(* Logix 5000 project; controller SmartManufacturingCell Emulate 5570 rev 33.11; software revision 33.03; part 3 of 5 *)
(* tags used below, declared in another part *)
   ClearCell_CommandsReleased : BOOL;
   ClearCell_EquipmentReady : BOOL;
   ClearCellRequestONS : BOOL;
   Exit_ReadyForIndex : BOOL;
   Filling_ReadyForIndex : BOOL;
   Index_CommandsReleased : BOOL;
   Index_EquipmentReady : BOOL;
   IndexConfirmTimeout : TIMER;   // Non-retentive timer; preset in milliseconds.
   IndexTimeout : TIMER;   // Non-retentive timer; preset in milliseconds.
   Inspection_ReadyForIndex : BOOL;
   Production_CycleHealthy : BOOL;
   Production_ResetAllowed : BOOL;
   Production_ResetCommandsReleased : BOOL;
   Production_SensorsClear : BOOL;
   Production_TrackingEmpty : BOOL;
   ProductionResetONS : BOOL;
   TrackingMismatchDelay : TIMER;   // Non-retentive timer; preset in milliseconds.
   Conveyor_Flt_FailToStart : BOOL;   // Conveyor commanded but running feedback missing for 2 s Latched; clear cell, remove cause, then fresh Reset.
   Exit_Flt_DischargeTimeout : BOOL;   // Good or reject bottle departure not confirmed within 3 s Latched; clear cell, remove cause, then fresh Reset.
   Exit_Sts_State : DINT;   // 0 Empty; 10 Waiting; 20 Good discharge; 30 Extending; 40 Reject discharge; 50 Retracting; 60 Complete; 90 Faulted
   Filling_Flt_FillTimeout : BOOL;   // Fill completion not received within 4 s Latched; clear cell, remove cause, then fresh Reset.
   Filling_Flt_ValveFailToClose : BOOL;   // Fill valve did not close within 2 s Latched; clear cell, remove cause, then fresh Reset.
   Filling_Sts_State : DINT;   // 0 Empty; 10 Waiting; 20 Filling; 30 Closing; 40 Complete; 90 Faulted
   HMI_Cmd_ClearCell : BOOL;   // Request removal of simulated bottles during fault recovery
   HMI_Cmd_ConveyorJog : BOOL;   // Request conveyor movement while held
   HMI_Cmd_FillValveOpen : BOOL;
   HMI_Cmd_LoadBottle : BOOL;   // Request one simulated bottle at the available entry position
   HMI_Cmd_RejectExtend : BOOL;
   HMI_Cmd_Reset : BOOL;   // Request fault reset after recovery conditions are satisfied
   HMI_Cmd_Start : BOOL;   // Request automatic production start
   HMI_Cmd_Stop : BOOL;   // Request controlled production stop
   Inspection_Flt_Timeout : BOOL;   // Inspection did not finish within 3 s Latched; clear cell, remove cause, then fresh Reset.
   Inspection_Sts_State : DINT;   // 0 Empty; 10 Waiting; 20 Inspecting; 40 Complete; 90 Faulted
   Production_Bottles : UDT_Bottle[4];
   Production_Flt_IndexConfirmTimeout : BOOL;   // Post-index positions not confirmed within 1 s Latched; clear cell, remove cause, then fresh Reset.
   Production_Flt_IndexInterlock : BOOL;   // Movement interlock lost during indexing Latched; clear cell, remove cause, then fresh Reset.
   Production_Flt_IndexTimeout : BOOL;   // Index completion not received within 3 s Latched; clear cell, remove cause, then fresh Reset.
   Production_Flt_InvalidConfiguration : BOOL;   // Fill or inspection time outside permitted limits Latched; clear cell, remove cause, then fresh Reset.
   Production_Flt_InvalidState : BOOL;   // Machine, sequence, station state, or mode combination invalid Latched; clear cell, remove cause, then fresh Reset.
   Production_Flt_StartupRecoveryRequired : BOOL;   // Restart found bottles or interrupted activity Latched; clear cell, remove cause, then fresh Reset.
   Production_Flt_TrackingMismatch : BOOL;   // Stationary bottle tracking and sensors disagree or processing history invalid Latched; clear cell, remove cause, then fr
   Production_Stats_RecoveryLossCount : DINT;   // Retained RecoveryLossCount; count only confirmed departures (recovery losses separate).
   Production_Sts_ClearCellAccepted : BOOL;
   Production_Sts_ClearCellAllowed : BOOL;
   Production_Sts_IndexAllowed : BOOL;
   Production_Sts_IndexCommitted : BOOL;   // Bottle records transferred for the current confirmed index; cleared outside ConfirmPositions.
   Production_Sts_IndexDemand : BOOL;
   Production_Sts_IndexPositionsMatch : BOOL;   // Post-index positions verified in ConfirmPositions with conveyor stopped.
   Production_Sts_LoadAccepted : BOOL;
   Production_Sts_ResetAccepted : BOOL;
   Production_Sts_SequenceState : DINT;   // 0 = Idle 10 = ProcessStations 20 = Indexing 30 = ConfirmPositions
   Production_Sts_StationsReady : BOOL;
   Reject_Flt_FailToExtend : BOOL;   // Reject actuator did not extend within 2 s Latched; clear cell, remove cause, then fresh Reset.
   Reject_Flt_FailToRetract : BOOL;   // Reject actuator did not retract within 2 s Latched; clear cell, remove cause, then fresh Reset.
   Sim_In_ConveyorRunning : BOOL;   // Simulated conveyor movement feedback
   Sim_In_EntryPE : BOOL;   // Simulated bottle detected at entry
   Sim_In_ExitPE : BOOL;   // Simulated bottle detected at Reject/Exit position
   Sim_In_FillPE : BOOL;   // Simulated bottle detected at filling position
   Sim_In_FillValveClosed : BOOL;   // Simulated fill valve confirmed closed
   Sim_In_GoodExitPE : BOOL;   // Bottle detected passing through good discharge path
   Sim_In_IndexComplete : BOOL;   // Simulated conveyor completed one station-spacing movement
   Sim_In_InspectionPE : BOOL;   // Simulated bottle detected at inspection position
   Sim_In_RejectExitPE : BOOL;   // Bottle detected passing through reject discharge path
   Sim_In_RejectExtended : BOOL;   // Simulated reject actuator confirmed extended
   Sim_In_RejectRetracted : BOOL;   // Simulated reject actuator confirmed retracted
   Sim_Out_ConveyorRun : BOOL;   // Command simulated conveyor to run
   Sim_Out_FillValveOpen : BOOL;   // Command simulated fill valve to open
   Sim_Out_GoodDischargeRun : BOOL;   // Command simulated good-bottle discharge mechanism to run
   Sim_Out_RejectExtend : BOOL;   // Command simulated reject actuator to extend
   Sys_Sts_AutoMode : BOOL;   // Auto mode accepted and active
   Sys_Sts_BlockingFault : BOOL;   // Active blocking fault prevents production and manual equipment operation.
   Sys_Sts_MachineState : DINT;   // 0 = Stopped 10 = Running 20 = Stopping 30 = Faulted
   Sys_Sts_ManualMode : BOOL;   // Manual mode accepted and active
   Sys_Sts_ResetAllowed : BOOL;   // Sys Sts ResetAllowed
   Sys_Sts_StartupReady : BOOL;   // Sys Sts StartupReady
(* Program_Production, continued *)

ROUTINE Bottle_Tracking   (* structured text *)
   if Production_Sts_SequenceState <> 30 then
   	Production_Sts_IndexCommitted := 0;
   elsif Production_Sts_IndexPositionsMatch AND NOT Production_Sts_IndexCommitted then
   
   	// Copy downstream first to preserve seach source record.
   	COP(Production_Bottles[2], Production_Bottles[3], 1);
   	COP(Production_Bottles[1], Production_Bottles[2], 1);
   	COP(Production_Bottles[0], Production_Bottles[1], 1);
   
    	// Entry is empty after the confirmed movement.
       Production_Bottles[0].Occupied := 0;
       Production_Bottles[0].FillComplete := 0;
       Production_Bottles[0].InspectionComplete := 0;
       Production_Bottles[0].RejectRequired := 0;
   
       Production_Sts_IndexCommitted := 1;
   end_if;
END_ROUTINE

ROUTINE Clear_Cell   (* ladder *)
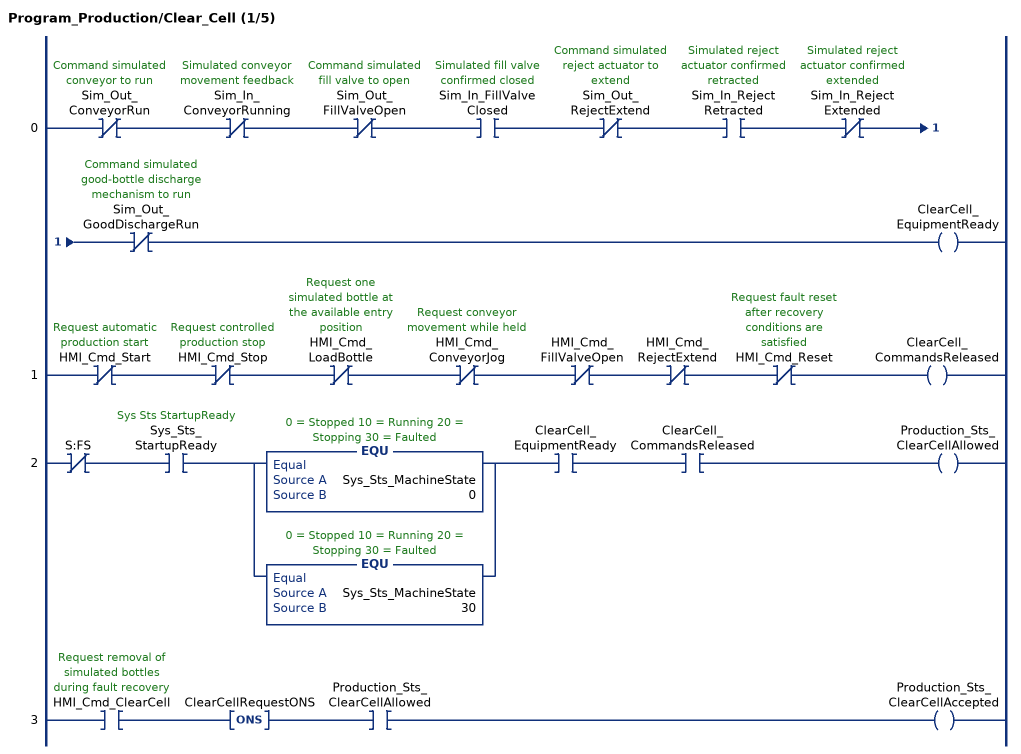
   0: XIO(Sim_Out_ConveyorRun)XIO(Sim_In_ConveyorRunning)XIO(Sim_Out_FillValveOpen)XIC(Sim_In_FillValveClosed)XIO(Sim_Out_RejectExtend)XIC(Sim_In_RejectRetracted)XIO(Sim_In_RejectExtended)XIO(Sim_Out_GoodDischargeRun)OTE(ClearCell_EquipmentReady);
   1: XIO(HMI_Cmd_Start)XIO(HMI_Cmd_Stop)XIO(HMI_Cmd_LoadBottle)XIO(HMI_Cmd_ConveyorJog)XIO(HMI_Cmd_FillValveOpen)XIO(HMI_Cmd_RejectExtend)XIO(HMI_Cmd_Reset)OTE(ClearCell_CommandsReleased);
   2: XIO(S:FS)XIC(Sys_Sts_StartupReady)[EQU(Sys_Sts_MachineState,0) ,EQU(Sys_Sts_MachineState,30) ]XIC(ClearCell_EquipmentReady)XIC(ClearCell_CommandsReleased)OTE(Production_Sts_ClearCellAllowed);
   3: XIC(HMI_Cmd_ClearCell)ONS(ClearCellRequestONS)XIC(Production_Sts_ClearCellAllowed)OTE(Production_Sts_ClearCellAccepted);
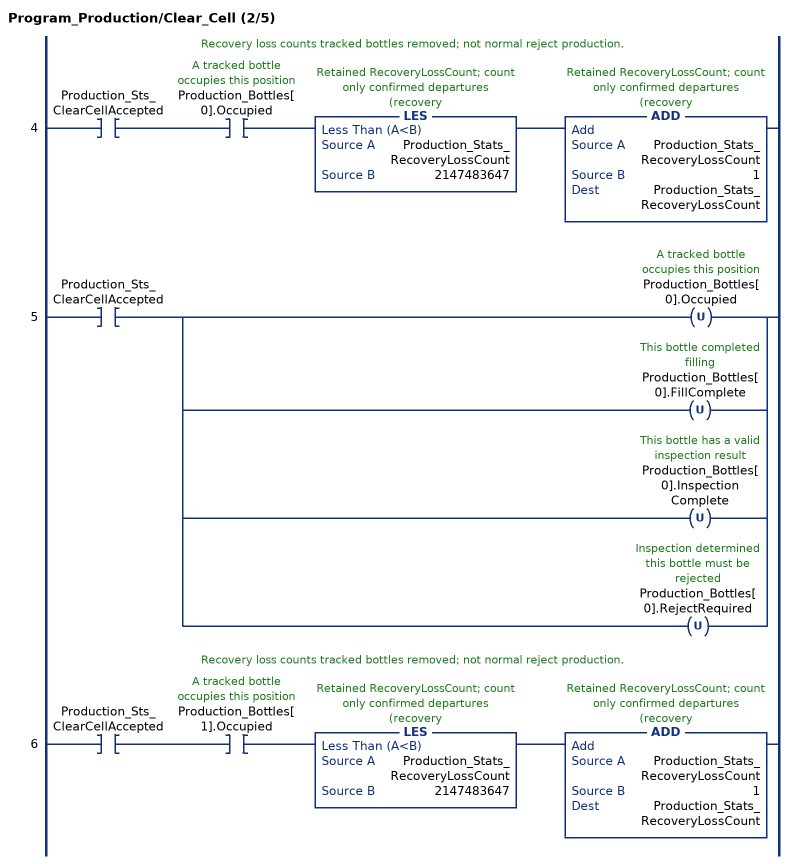
   // Recovery loss counts tracked bottles removed; not normal reject production.
   4: XIC(Production_Sts_ClearCellAccepted)XIC(Production_Bottles[0].Occupied)LES(Production_Stats_RecoveryLossCount,2147483647)ADD(Production_Stats_RecoveryLossCount,1,Production_Stats_RecoveryLossCount);
   5: XIC(Production_Sts_ClearCellAccepted)[OTU(Production_Bottles[0].Occupied) ,OTU(Production_Bottles[0].FillComplete) ,OTU(Production_Bottles[0].InspectionComplete) ,OTU(Production_Bottles[0].RejectRequired) ];
   // Recovery loss counts tracked bottles removed; not normal reject production.
   6: XIC(Production_Sts_ClearCellAccepted)XIC(Production_Bottles[1].Occupied)LES(Production_Stats_RecoveryLossCount,2147483647)ADD(Production_Stats_RecoveryLossCount,1,Production_Stats_RecoveryLossCount);
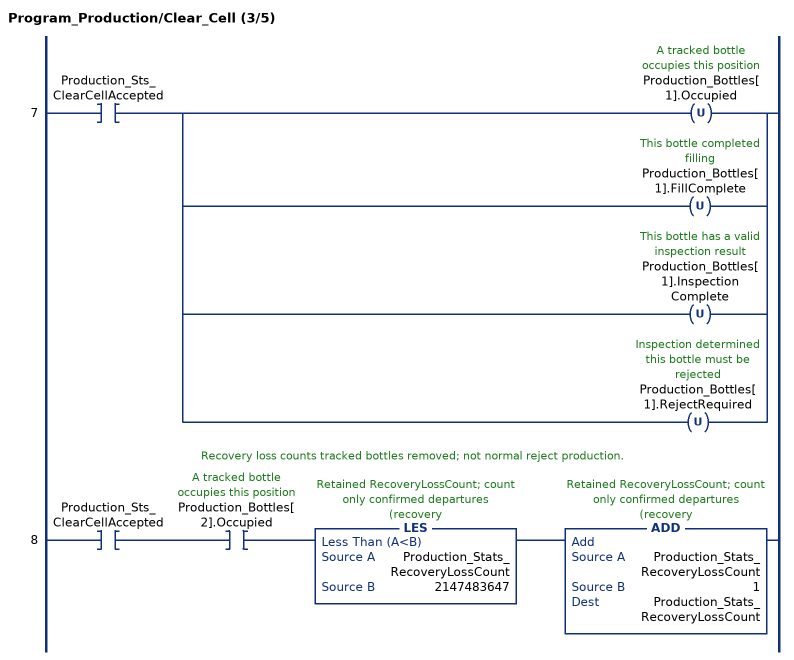
   7: XIC(Production_Sts_ClearCellAccepted)[OTU(Production_Bottles[1].Occupied) ,OTU(Production_Bottles[1].FillComplete) ,OTU(Production_Bottles[1].InspectionComplete) ,OTU(Production_Bottles[1].RejectRequired) ];
   // Recovery loss counts tracked bottles removed; not normal reject production.
   8: XIC(Production_Sts_ClearCellAccepted)XIC(Production_Bottles[2].Occupied)LES(Production_Stats_RecoveryLossCount,2147483647)ADD(Production_Stats_RecoveryLossCount,1,Production_Stats_RecoveryLossCount);
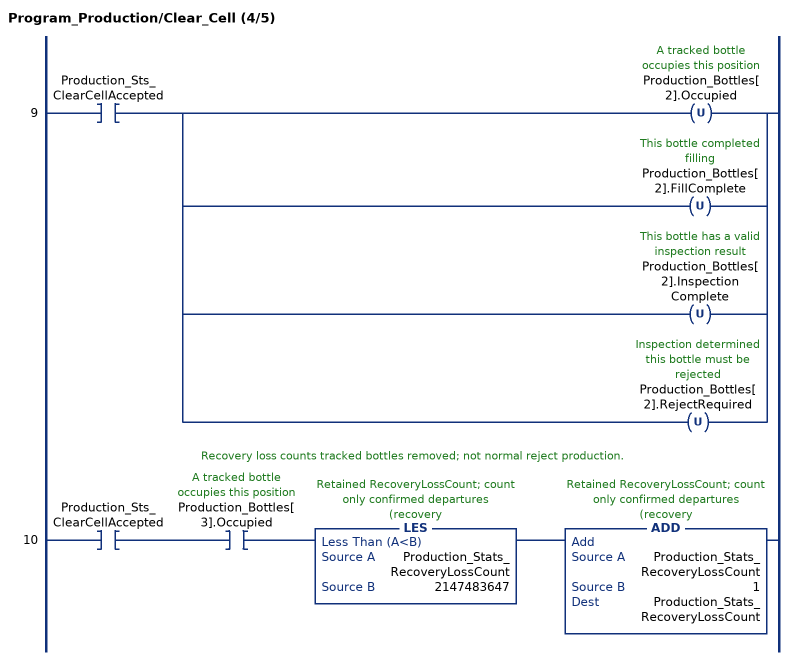
   9: XIC(Production_Sts_ClearCellAccepted)[OTU(Production_Bottles[2].Occupied) ,OTU(Production_Bottles[2].FillComplete) ,OTU(Production_Bottles[2].InspectionComplete) ,OTU(Production_Bottles[2].RejectRequired) ];
   // Recovery loss counts tracked bottles removed; not normal reject production.
   10: XIC(Production_Sts_ClearCellAccepted)XIC(Production_Bottles[3].Occupied)LES(Production_Stats_RecoveryLossCount,2147483647)ADD(Production_Stats_RecoveryLossCount,1,Production_Stats_RecoveryLossCount);
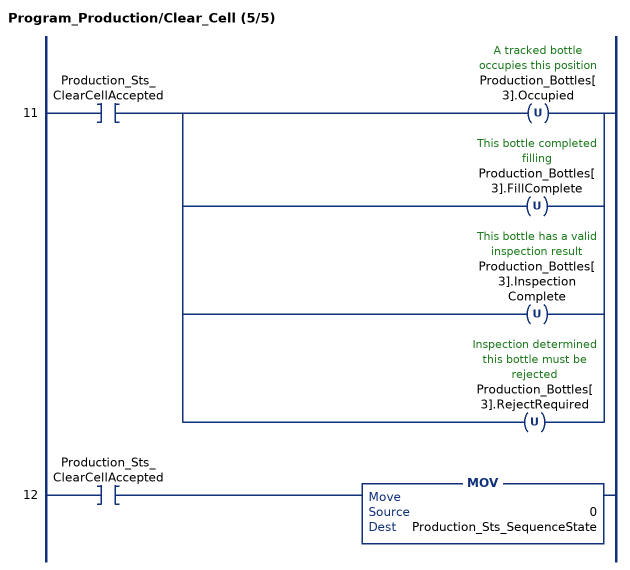
   11: XIC(Production_Sts_ClearCellAccepted)[OTU(Production_Bottles[3].Occupied) ,OTU(Production_Bottles[3].FillComplete) ,OTU(Production_Bottles[3].InspectionComplete) ,OTU(Production_Bottles[3].RejectRequired) ];
   12: XIC(Production_Sts_ClearCellAccepted)MOV(0,Production_Sts_SequenceState);
END_ROUTINE

ROUTINE Index_Confirmation   (* structured text *)
   Production_Sts_IndexPositionsMatch :=
       (Production_Sts_SequenceState = 30)
       AND (
           (Sys_Sts_MachineState = 10)
           OR (Sys_Sts_MachineState = 20)
       )
       AND Sys_Sts_AutoMode
       AND NOT Sys_Sts_ManualMode
       AND NOT Sys_Sts_BlockingFault
       AND NOT Sim_Out_ConveyorRun
       AND NOT Sim_In_ConveyorRunning
       AND NOT Production_Bottles[3].Occupied
       AND NOT Sim_In_EntryPE
       AND NOT (Sim_In_FillPE XOR Production_Bottles[0].Occupied)
       AND NOT (Sim_In_InspectionPE XOR Production_Bottles[1].Occupied)
       AND NOT (Sim_In_ExitPE XOR Production_Bottles[2].Occupied);
END_ROUTINE

ROUTINE Index_Permissives   (* ladder *)
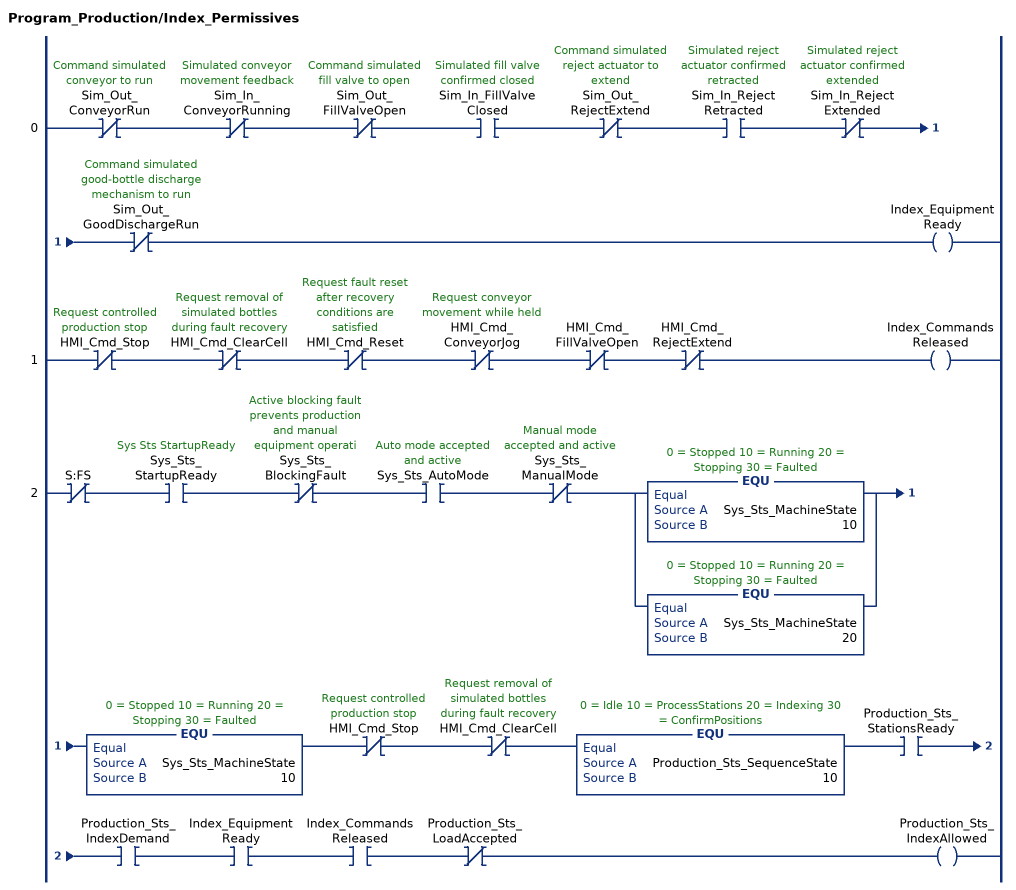
   0: XIO(Sim_Out_ConveyorRun)XIO(Sim_In_ConveyorRunning)XIO(Sim_Out_FillValveOpen)XIC(Sim_In_FillValveClosed)XIO(Sim_Out_RejectExtend)XIC(Sim_In_RejectRetracted)XIO(Sim_In_RejectExtended)XIO(Sim_Out_GoodDischargeRun)OTE(Index_EquipmentReady);
   1: XIO(HMI_Cmd_Stop)XIO(HMI_Cmd_ClearCell)XIO(HMI_Cmd_Reset)XIO(HMI_Cmd_ConveyorJog)XIO(HMI_Cmd_FillValveOpen)XIO(HMI_Cmd_RejectExtend)OTE(Index_CommandsReleased);
   2: XIO(S:FS)XIC(Sys_Sts_StartupReady)XIO(Sys_Sts_BlockingFault)XIC(Sys_Sts_AutoMode)XIO(Sys_Sts_ManualMode)[EQU(Sys_Sts_MachineState,10) ,EQU(Sys_Sts_MachineState,20) ]EQU(Sys_Sts_MachineState,10)XIO(HMI_Cmd_Stop)XIO(HMI_Cmd_ClearCell)EQU(Production_Sts_SequenceState,10)XIC(Production_Sts_StationsReady)XIC(Production_Sts_IndexDemand)XIC(Index_EquipmentReady)XIC(Index_CommandsReleased)XIO(Production_Sts_LoadAccepted)OTE(Production_Sts_IndexAllowed);
END_ROUTINE

ROUTINE Index_Readiness   (* ladder *)
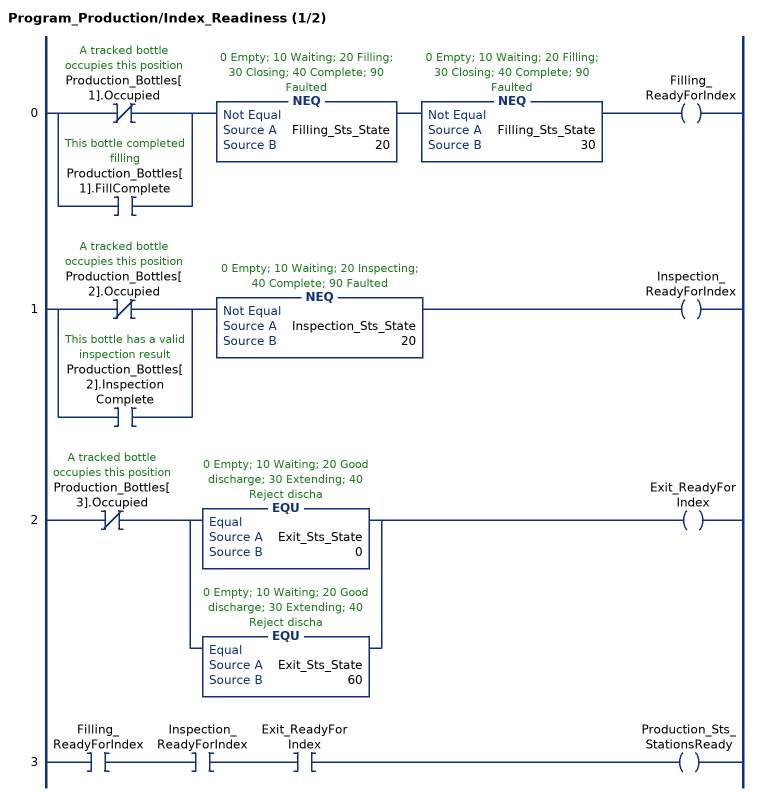
   0: [XIO(Production_Bottles[1].Occupied) ,XIC(Production_Bottles[1].FillComplete) ]NEQ(Filling_Sts_State,20)NEQ(Filling_Sts_State,30)OTE(Filling_ReadyForIndex);
   1: [XIO(Production_Bottles[2].Occupied) ,XIC(Production_Bottles[2].InspectionComplete) ]NEQ(Inspection_Sts_State,20)OTE(Inspection_ReadyForIndex);
   2: XIO(Production_Bottles[3].Occupied)[EQU(Exit_Sts_State,0) ,EQU(Exit_Sts_State,60) ]OTE(Exit_ReadyForIndex);
   3: XIC(Filling_ReadyForIndex)XIC(Inspection_ReadyForIndex)XIC(Exit_ReadyForIndex)OTE(Production_Sts_StationsReady);
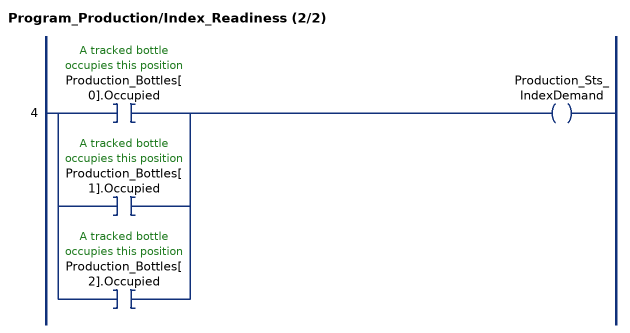
   4: [XIC(Production_Bottles[0].Occupied) ,XIC(Production_Bottles[1].Occupied) ,XIC(Production_Bottles[2].Occupied) ]OTE(Production_Sts_IndexDemand);
END_ROUTINE

ROUTINE MainRoutine   (* ladder *)
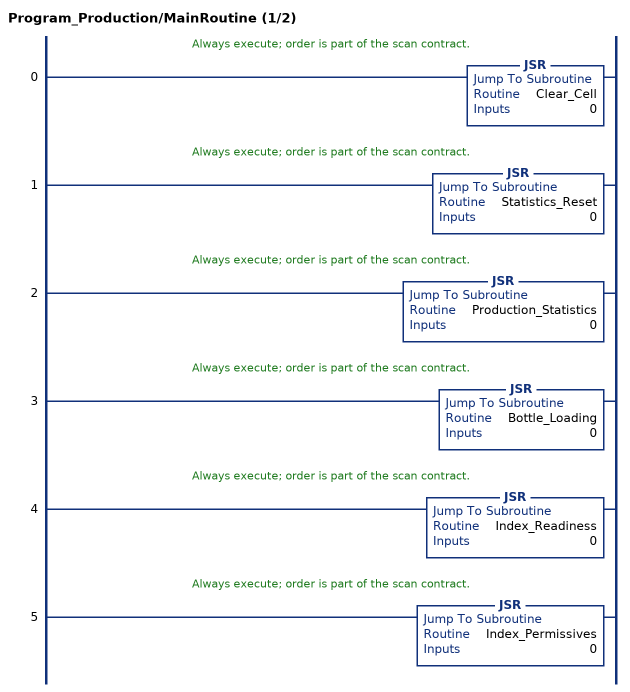
   // Always execute; order is part of the scan contract.
   0: JSR(Clear_Cell,0);
   // Always execute; order is part of the scan contract.
   1: JSR(Statistics_Reset,0);
   // Always execute; order is part of the scan contract.
   2: JSR(Production_Statistics,0);
   // Always execute; order is part of the scan contract.
   3: JSR(Bottle_Loading,0);
   // Always execute; order is part of the scan contract.
   4: JSR(Index_Readiness,0);
   // Always execute; order is part of the scan contract.
   5: JSR(Index_Permissives,0);
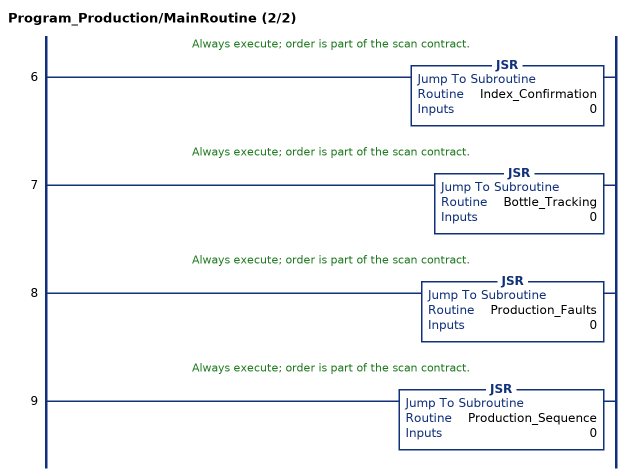
   // Always execute; order is part of the scan contract.
   6: JSR(Index_Confirmation,0);
   // Always execute; order is part of the scan contract.
   7: JSR(Bottle_Tracking,0);
   // Always execute; order is part of the scan contract.
   8: JSR(Production_Faults,0);
   // Always execute; order is part of the scan contract.
   9: JSR(Production_Sequence,0);
END_ROUTINE

ROUTINE Production_Faults   (* ladder *)
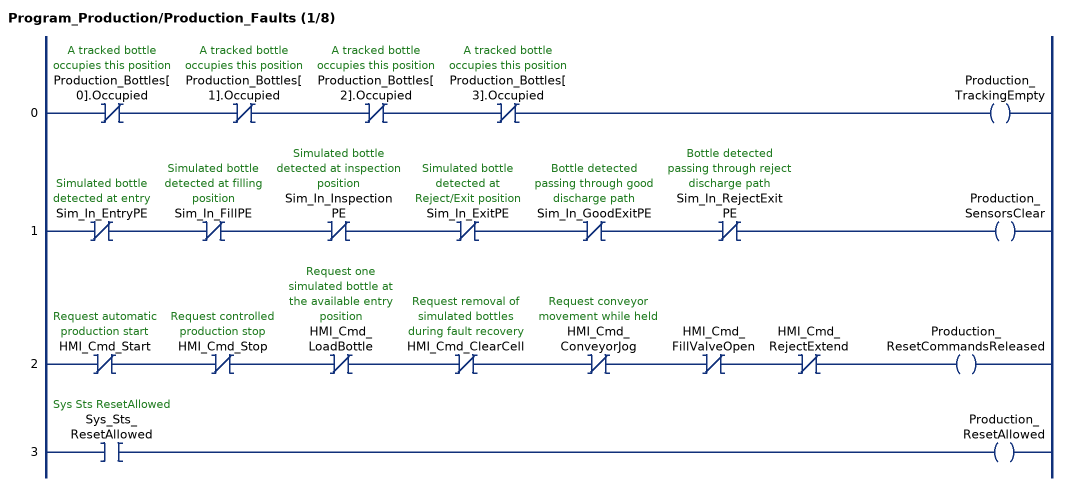
   0: XIO(Production_Bottles[0].Occupied)XIO(Production_Bottles[1].Occupied)XIO(Production_Bottles[2].Occupied)XIO(Production_Bottles[3].Occupied)OTE(Production_TrackingEmpty);
   1: XIO(Sim_In_EntryPE)XIO(Sim_In_FillPE)XIO(Sim_In_InspectionPE)XIO(Sim_In_ExitPE)XIO(Sim_In_GoodExitPE)XIO(Sim_In_RejectExitPE)OTE(Production_SensorsClear);
   2: XIO(HMI_Cmd_Start)XIO(HMI_Cmd_Stop)XIO(HMI_Cmd_LoadBottle)XIO(HMI_Cmd_ClearCell)XIO(HMI_Cmd_ConveyorJog)XIO(HMI_Cmd_FillValveOpen)XIO(HMI_Cmd_RejectExtend)OTE(Production_ResetCommandsReleased);
   3: XIC(Sys_Sts_ResetAllowed)OTE(Production_ResetAllowed);
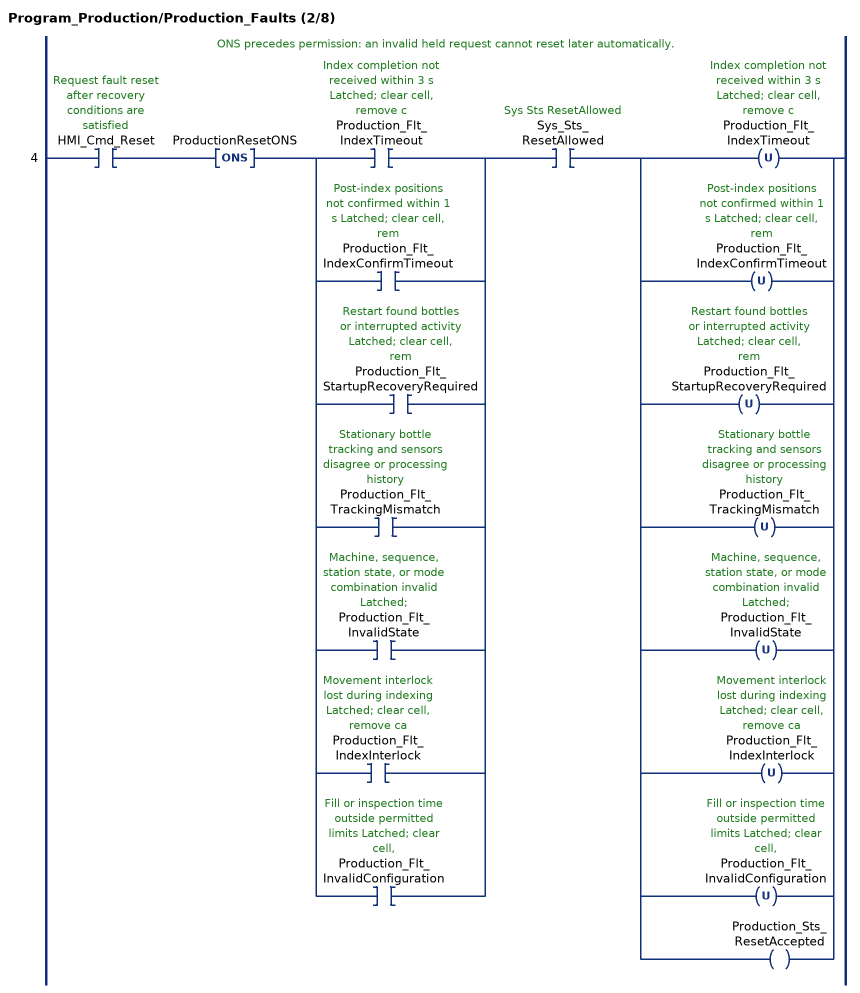
   // ONS precedes permission: an invalid held request cannot reset later automatically.
   4: XIC(HMI_Cmd_Reset)ONS(ProductionResetONS)[XIC(Production_Flt_IndexTimeout) ,XIC(Production_Flt_IndexConfirmTimeout) ,XIC(Production_Flt_StartupRecoveryRequired) ,XIC(Production_Flt_TrackingMismatch) ,XIC(Production_Flt_InvalidState) ,XIC(Production_Flt_IndexInterlock) ,XIC(Production_Flt_InvalidConfiguration) ]XIC(Sys_Sts_ResetAllowed)[OTU(Production_Flt_IndexTimeout) ,OTU(Production_Flt_IndexConfirmTimeout) ,OTU(Production_Flt_StartupRecoveryRequired) ,OTU(Production_Flt_TrackingMismatch) ,OTU(Production_Flt_InvalidState) ,OTU(Production_Flt_IndexInterlock) ,OTU(Production_Flt_InvalidConfiguration) ,OTE(Production_Sts_ResetAccepted) ];
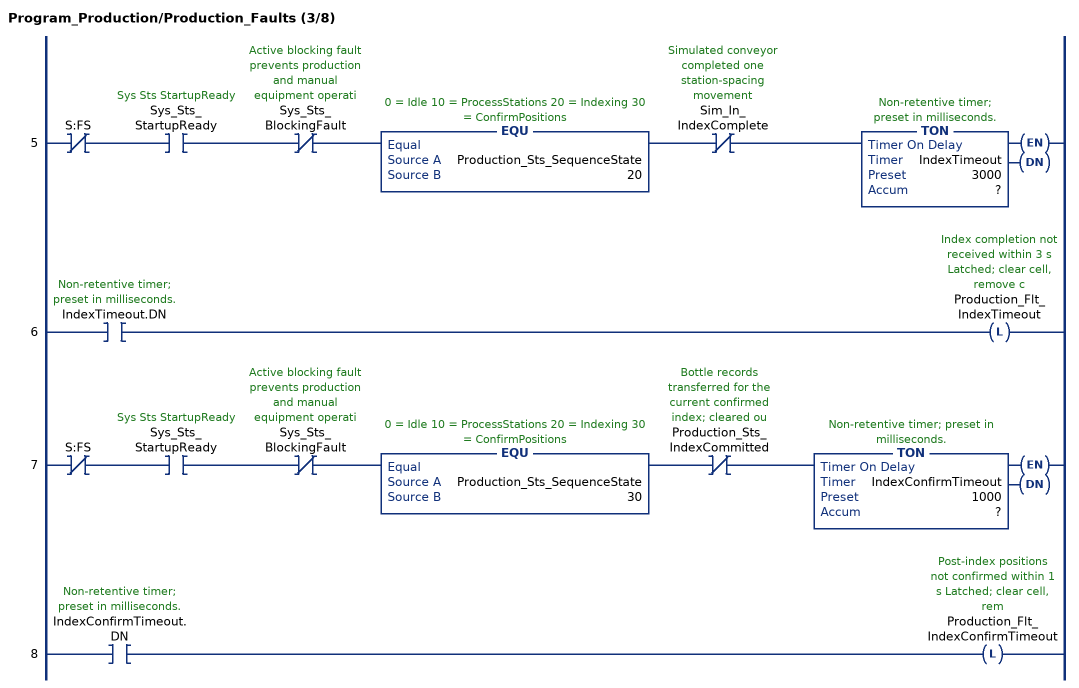
   5: XIO(S:FS)XIC(Sys_Sts_StartupReady)XIO(Sys_Sts_BlockingFault)EQU(Production_Sts_SequenceState,20)XIO(Sim_In_IndexComplete)TON(IndexTimeout,?,?);
   6: XIC(IndexTimeout.DN)OTL(Production_Flt_IndexTimeout);
   7: XIO(S:FS)XIC(Sys_Sts_StartupReady)XIO(Sys_Sts_BlockingFault)EQU(Production_Sts_SequenceState,30)XIO(Production_Sts_IndexCommitted)TON(IndexConfirmTimeout,?,?);
   8: XIC(IndexConfirmTimeout.DN)OTL(Production_Flt_IndexConfirmTimeout);
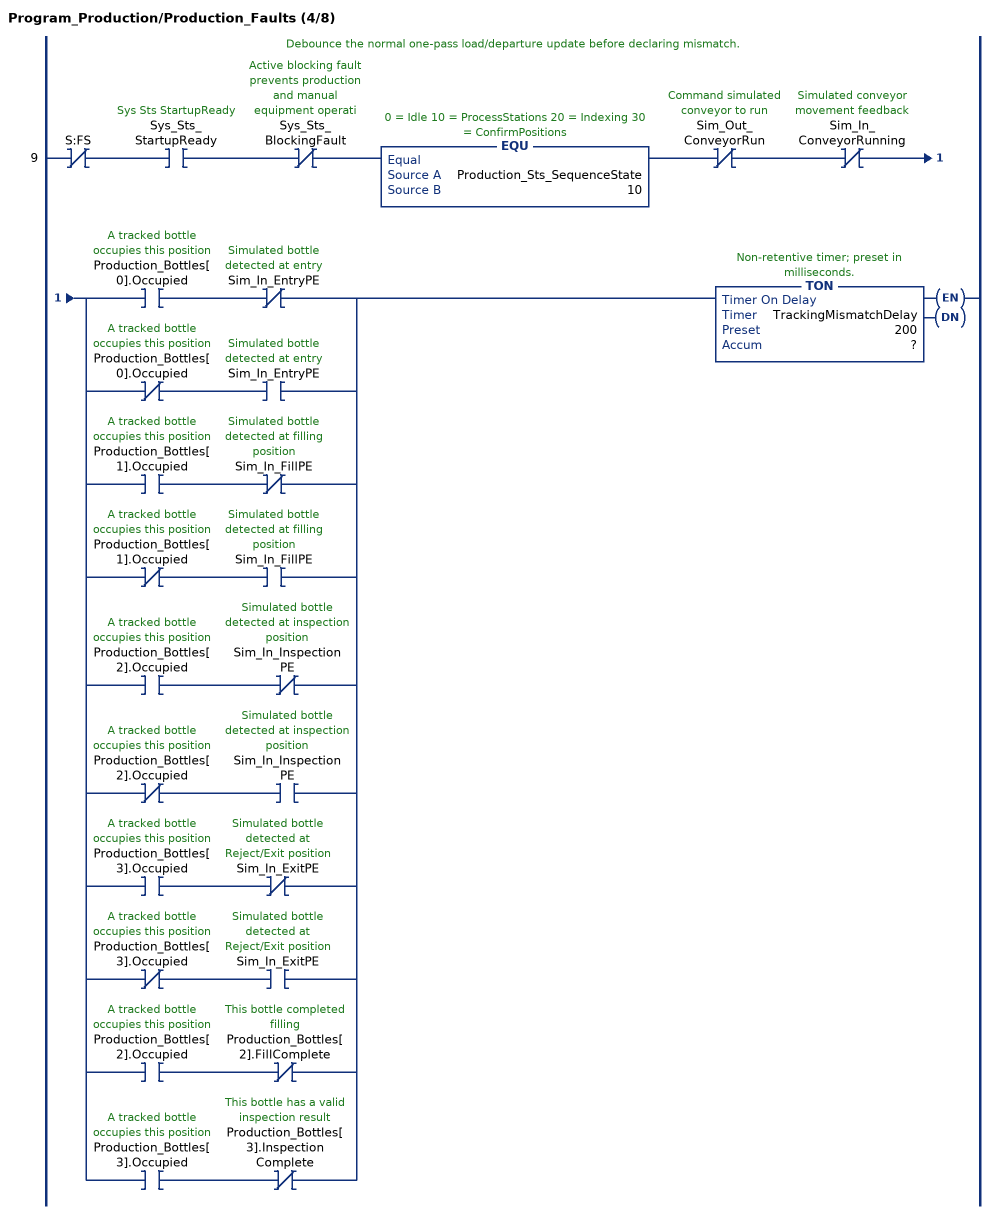
   // Debounce the normal one-pass load/departure update before declaring mismatch.
   9: XIO(S:FS)XIC(Sys_Sts_StartupReady)XIO(Sys_Sts_BlockingFault)EQU(Production_Sts_SequenceState,10)XIO(Sim_Out_ConveyorRun)XIO(Sim_In_ConveyorRunning)[[XIC(Production_Bottles[0].Occupied) XIO(Sim_In_EntryPE) ,XIO(Production_Bottles[0].Occupied) XIC(Sim_In_EntryPE) ] ,[XIC(Production_Bottles[1].Occupied) XIO(Sim_In_FillPE) ,XIO(Production_Bottles[1].Occupied) XIC(Sim_In_FillPE) ] ,[XIC(Production_Bottles[2].Occupied) XIO(Sim_In_InspectionPE) ,XIO(Production_Bottles[2].Occupied) XIC(Sim_In_InspectionPE) ] ,[XIC(Production_Bottles[3].Occupied) XIO(Sim_In_ExitPE) ,XIO(Production_Bottles[3].Occupied) XIC(Sim_In_ExitPE) ] ,XIC(Production_Bottles[2].Occupied) XIO(Production_Bottles[2].FillComplete) ,XIC(Production_Bottles[3].Occupied) XIO(Production_Bottles[3].InspectionComplete) ]TON(TrackingMismatchDelay,?,?);
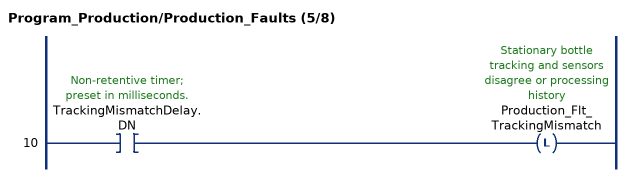
   10: XIC(TrackingMismatchDelay.DN)OTL(Production_Flt_TrackingMismatch);
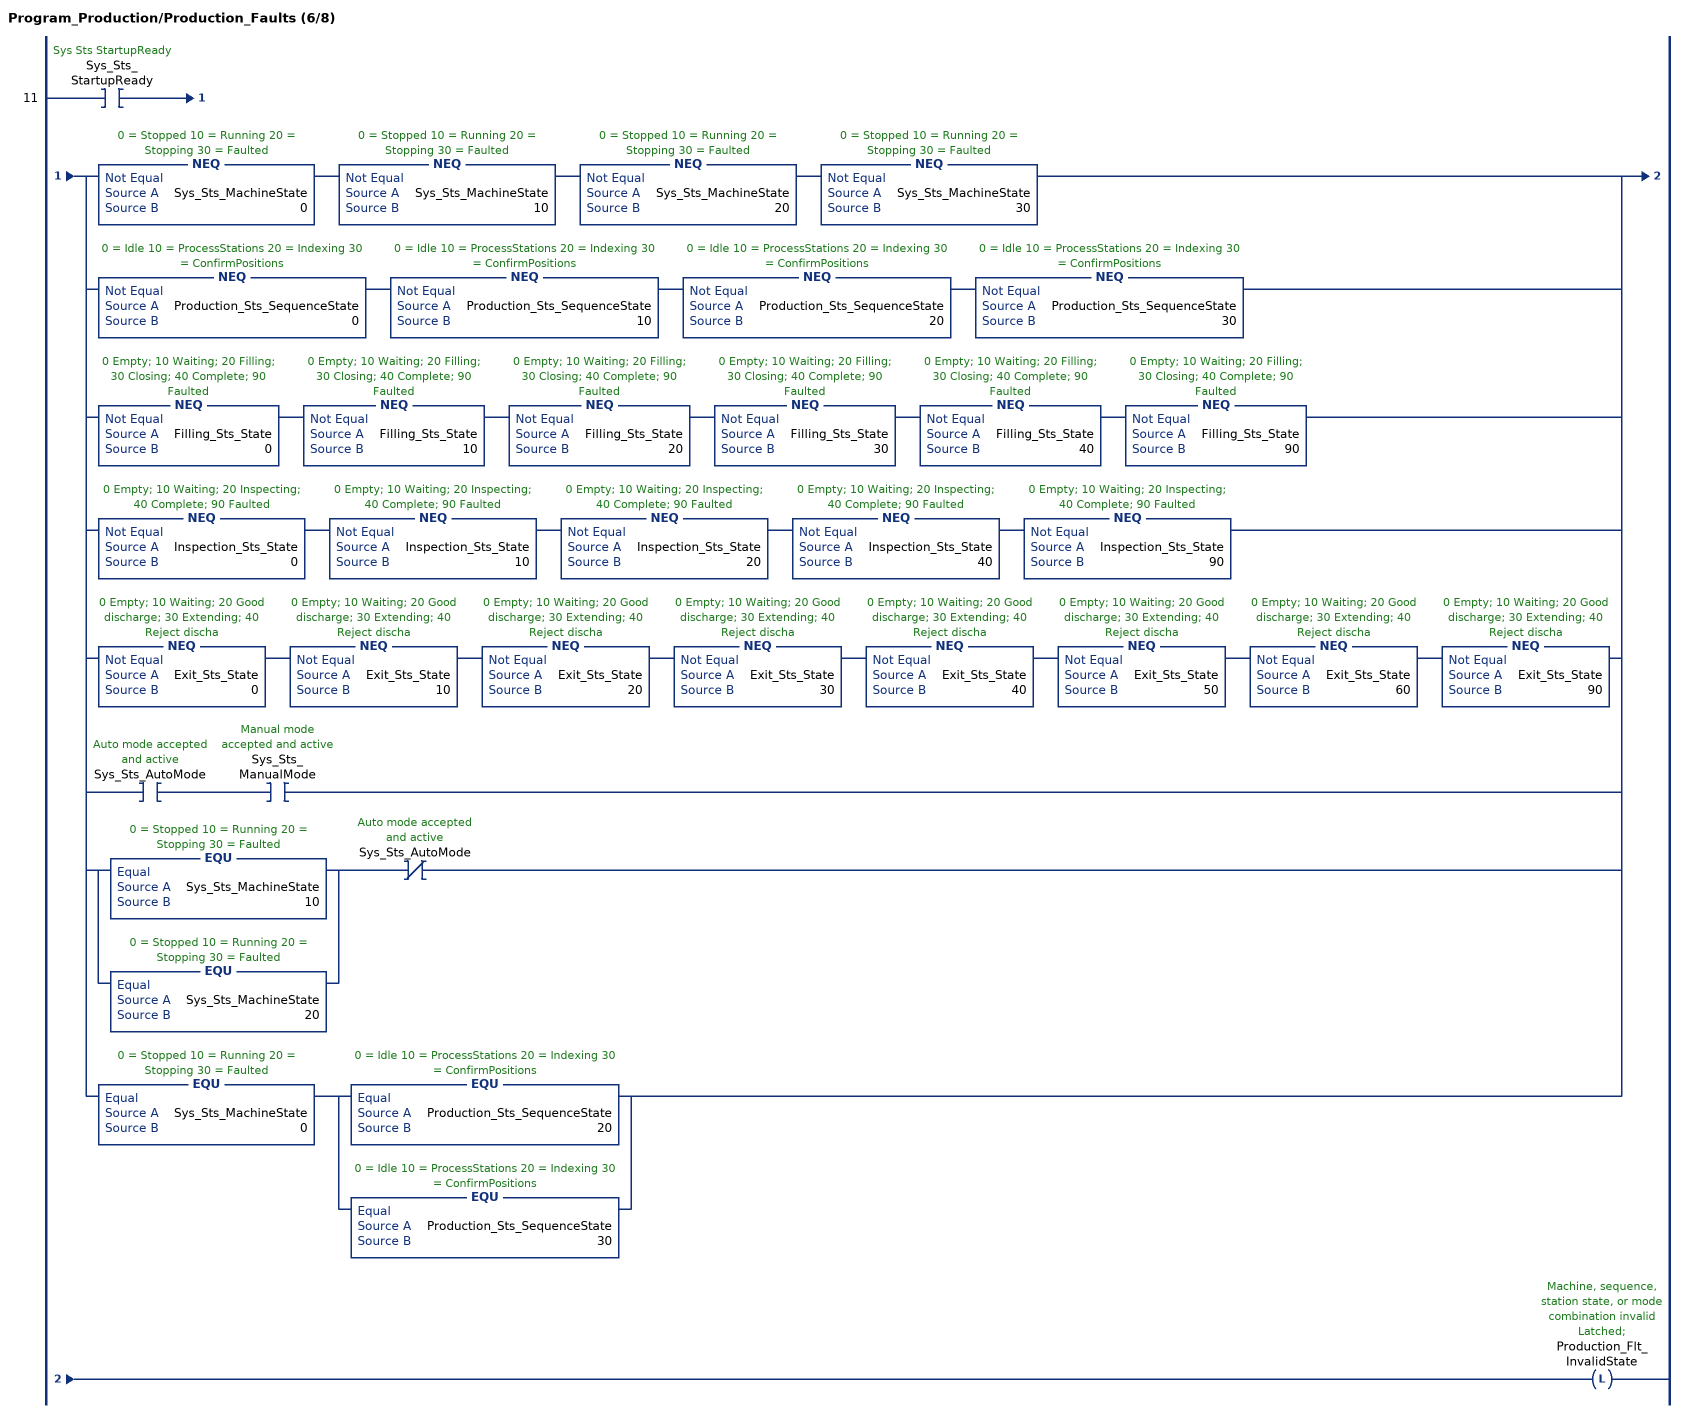
   11: XIC(Sys_Sts_StartupReady)[NEQ(Sys_Sts_MachineState,0) NEQ(Sys_Sts_MachineState,10) NEQ(Sys_Sts_MachineState,20) NEQ(Sys_Sts_MachineState,30) ,NEQ(Production_Sts_SequenceState,0) NEQ(Production_Sts_SequenceState,10) NEQ(Production_Sts_SequenceState,20) NEQ(Production_Sts_SequenceState,30) ,NEQ(Filling_Sts_State,0) NEQ(Filling_Sts_State,10) NEQ(Filling_Sts_State,20) NEQ(Filling_Sts_State,30) NEQ(Filling_Sts_State,40) NEQ(Filling_Sts_State,90) ,NEQ(Inspection_Sts_State,0) NEQ(Inspection_Sts_State,10) NEQ(Inspection_Sts_State,20) NEQ(Inspection_Sts_State,40) NEQ(Inspection_Sts_State,90) ,NEQ(Exit_Sts_State,0) NEQ(Exit_Sts_State,10) NEQ(Exit_Sts_State,20) NEQ(Exit_Sts_State,30) NEQ(Exit_Sts_State,40) NEQ(Exit_Sts_State,50) NEQ(Exit_Sts_State,60) NEQ(Exit_Sts_State,90) ,XIC(Sys_Sts_AutoMode) XIC(Sys_Sts_ManualMode) ,[EQU(Sys_Sts_MachineState,10) ,EQU(Sys_Sts_MachineState,20) ] XIO(Sys_Sts_AutoMode) ,EQU(Sys_Sts_MachineState,0) [EQU(Production_Sts_SequenceState,20) ,EQU(Production_Sts_SequenceState,30) ] ]OTL(Production_Flt_InvalidState);
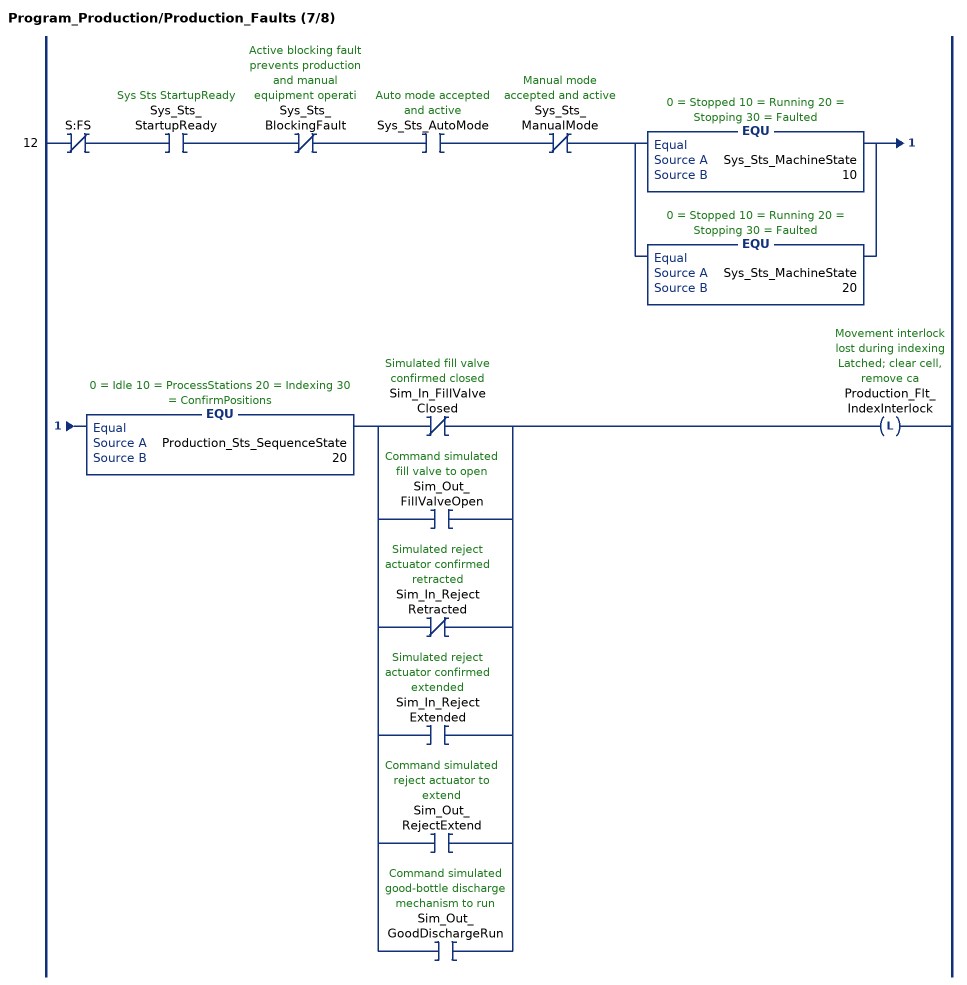
   12: XIO(S:FS)XIC(Sys_Sts_StartupReady)XIO(Sys_Sts_BlockingFault)XIC(Sys_Sts_AutoMode)XIO(Sys_Sts_ManualMode)[EQU(Sys_Sts_MachineState,10) ,EQU(Sys_Sts_MachineState,20) ]EQU(Production_Sts_SequenceState,20)[XIO(Sim_In_FillValveClosed) ,XIC(Sim_Out_FillValveOpen) ,XIO(Sim_In_RejectRetracted) ,XIC(Sim_In_RejectExtended) ,XIC(Sim_Out_RejectExtend) ,XIC(Sim_Out_GoodDischargeRun) ]OTL(Production_Flt_IndexInterlock);
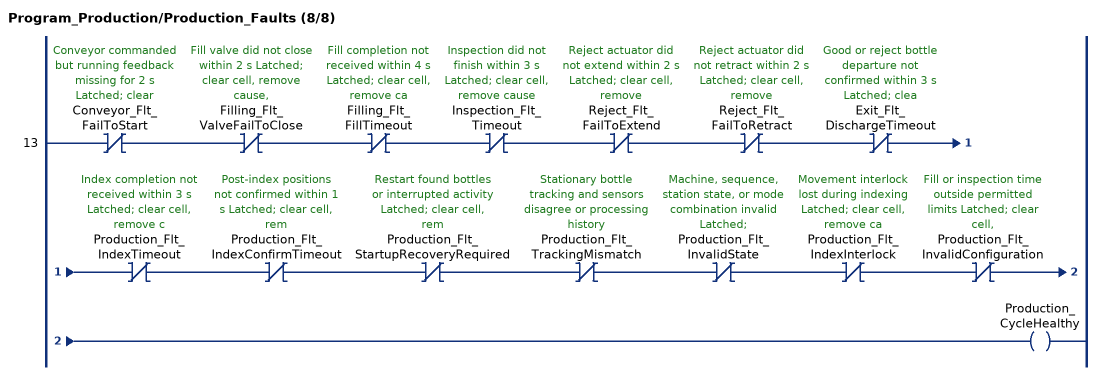
   13: XIO(Conveyor_Flt_FailToStart)XIO(Filling_Flt_ValveFailToClose)XIO(Filling_Flt_FillTimeout)XIO(Inspection_Flt_Timeout)XIO(Reject_Flt_FailToExtend)XIO(Reject_Flt_FailToRetract)XIO(Exit_Flt_DischargeTimeout)XIO(Production_Flt_IndexTimeout)XIO(Production_Flt_IndexConfirmTimeout)XIO(Production_Flt_StartupRecoveryRequired)XIO(Production_Flt_TrackingMismatch)XIO(Production_Flt_InvalidState)XIO(Production_Flt_IndexInterlock)XIO(Production_Flt_InvalidConfiguration)OTE(Production_CycleHealthy);
END_ROUTINE
